Fanuc KAREL source: ka00227.KL

PROGRAM KA00227
%STACKSIZE=65535
%PRIORITY=65535
%NOLOCKGROUP
-- UNRESOLVED DECLARATIONS (source type spelling not recovered)
-- SRC : TYPE_0x1100 (type_u16=0x1100)
-- DST : TYPE_0x1100 (type_u16=0x1100)
BEGIN
-- UNRESOLVED_PC line 7 opcodes [22 22 30] marker_code=0
END KA00227
